(* IEC 61131-3 sources: model-first-plc-agent-ai/results/T1-W-08, 2 files *)

(* ---- a1_code.st ---- *)
FUNCTION_BLOCK ConveyorRuntime
VAR_INPUT
    sensor_a : BOOL;
    sensor_b : BOOL;
END_VAR
VAR_OUTPUT
    conveyor : BOOL := FALSE;
END_VAR
VAR
    command_latch : RS;
END_VAR

(* Q1 initially FALSE represents initial step x0.
   Q1 TRUE represents step x1. *)
command_latch(
    S := sensor_a AND NOT sensor_b,
    R1 := sensor_b
);

conveyor := command_latch.Q1;

END_FUNCTION_BLOCK

PROGRAM Main
VAR
    SensorA AT %IX100.0 : BOOL;
    SensorB AT %IX100.1 : BOOL;
    Conveyor AT %QX100.0 : BOOL;
END_VAR
VAR
    controller : ConveyorRuntime;
END_VAR

controller(
    sensor_a := SensorA,
    sensor_b := SensorB
);

Conveyor := controller.conveyor;

END_PROGRAM

(* ---- a2_code.st ---- *)
FUNCTION_BLOCK ConveyorControl
VAR_INPUT
    sensor_a : BOOL;
    sensor_b : BOOL;
END_VAR
VAR_OUTPUT
    conveyor : BOOL;
END_VAR
VAR
    command_latch : RS;
END_VAR

command_latch(S := sensor_a, R1 := sensor_b);
conveyor := command_latch.Q1;

END_FUNCTION_BLOCK

PROGRAM Main
VAR
    sensor_a AT %IX100.0 : BOOL;
    sensor_b AT %IX100.1 : BOOL;
    conveyor AT %QX100.0 : BOOL;
END_VAR
VAR
    controller : ConveyorControl;
END_VAR

controller(
    sensor_a := sensor_a,
    sensor_b := sensor_b,
    conveyor => conveyor
);

END_PROGRAM
